(* IEC 61131-3 sources: plc-process-lib/tests/POUs/Suites/FB_ControlValve_Test, 43 files *)

(* ---- AutoSpNaNHoldsWithWarning.method.decl.st ---- *)
// Задание автоматики не число (NaN из Modbus/ПИД): выход удерживается, CV_WRN_SP_INVALID; конечное
// задание — снова к нему, предупреждение снято.
METHOD PRIVATE AutoSpNaNHoldsWithWarning
VAR
    fbTime   : FB_FakeTime;          // подменное время, старт 1 ч
    fbCv     : FB_ControlValve;      // клапан под тестом
    stCmd    : ST_ControlValveCmd;   // команды HMI
    stRetain : ST_DeviceRetain;      // режим Manual по умолчанию
    stCfg    : ST_ControlValveCfg;   // конфигурация (умолчания: 0…100 %, без рампы)
    uBits    : U_RealBits;           // NaN по битам
END_VAR

(* ---- AutoToManualBumpless.method.decl.st ---- *)
// Auto 70 %: задание Manual следит (70 %). Переход в Manual при задании автоматики 20 %: выход остаётся
// 70 %, xAutoActive = FALSE; задание оператора 60 % — рампа 5 %/с от 70 %: 65 % через 1 с.
METHOD PRIVATE AutoToManualBumpless
VAR
    fbTime   : FB_FakeTime;          // подменное время, старт 1 ч
    fbCv     : FB_ControlValve;      // клапан под тестом
    stCmd    : ST_ControlValveCmd;   // команды HMI
    stRetain : ST_DeviceRetain;      // режим Manual по умолчанию
    stCfg    : ST_ControlValveCfg;   // конфигурация (умолчания: 0…100 %, без рампы)
    iStep    : INT;                  // шаг цикла
END_VAR

(* ---- AutoToManualBumpless.method.impl.st ---- *)
coUnit.TEST('ControlValve_AutoToManual_Bumpless');

stRetain.eRemoteMode := E_DeviceMode.Auto;
fbCv.rPosSpAuto_pct := 70.0;
fbCv(itfTime := fbTime, stCmd := stCmd, stRetain := stRetain, stCfg := stCfg);
AssertEquals_REAL(Expected := 70.0, Actual := fbCv.rOut_pct, Delta := 0.0, Message := 'Auto 70 %');
AssertTrue(Condition := fbCv.xAutoActive, Message := 'xAutoActive');
AssertEquals_REAL(Expected := 70.0, Actual := stCmd.rPosSpMan_pct, Delta := 0.0,
                  Message := 'manual setpoint tracks in Auto');
stCfg.rRateUp_pctps := 5.0;
stCfg.rRateDown_pctps := 5.0;
stCmd.stCommon.xSetManual := TRUE;
fbCv.rPosSpAuto_pct := 20.0;
fbTime.Advance(tStep := T#100MS);
fbCv(itfTime := fbTime, stCmd := stCmd, stRetain := stRetain, stCfg := stCfg);
AssertTrue(Condition := fbCv.Mode = E_DeviceMode.Manual, Message := 'Manual');
AssertEquals_REAL(Expected := 70.0, Actual := fbCv.rOut_pct, Delta := 0.0, Message := 'no bump');
AssertFalse(Condition := fbCv.xAutoActive, Message := 'xAutoActive off in Manual');
stCmd.rPosSpMan_pct := 60.0;
FOR iStep := 1 TO 10 DO
    fbTime.Advance(tStep := T#100MS);
    fbCv(itfTime := fbTime, stCmd := stCmd, stRetain := stRetain, stCfg := stCfg);
END_FOR
// источник: tools/reference/valve_reference.py, сценарий cv_bumpless (70 -> 60, 5 %/s, 1.0 s)
AssertEquals_REAL(Expected := 65.0, Actual := fbCv.rOut_pct, Delta := 1.0E-4,
                  Message := 'ramp from 70 %: 65 % after 1 s');

coUnit.TEST_FINISHED();

(* ---- CfgChecksSetBits.method.decl.st ---- *)
// Каждая проверка CheckConfig даёт свой бит wCfgErr: пределы (min < 0, max > 100, min >= max), скорость
// (< 0, NaN), положение безопасности вне 0…100, рассогласование при подключённой ОС (допуск 0, tDev = 0;
// без ОС не проверяется), плотное закрытие (< 0, >= rOutMax), реакция на отказ вне перечисления,
// приоритет тревоги.
METHOD PRIVATE CfgChecksSetBits
VAR
    fbTime   : FB_FakeTime;          // подменное время, старт 1 ч
    fbCv     : FB_ControlValve;      // клапан под тестом
    stCmd    : ST_ControlValveCmd;   // команды HMI
    stRetain : ST_DeviceRetain;      // режим Manual по умолчанию
    stCfg    : ST_ControlValveCfg;   // конфигурация (умолчания: 0…100 %, без рампы)
    uBad     : U_TestValveEnum;      // значение вне перечисления
    uBits    : U_RealBits;           // NaN по битам
    stSlot   : ST_AlarmCfg;          // копия слота тревоги
END_VAR

(* ---- DefaultCfgPassesCheck.method.decl.st ---- *)
// Умолчания ST_ControlValveCfg проходят CheckConfig; тип ControlValve, слотов тревог 4, приоритеты по
// умолчанию (PositionerFault — Medium, InterlockAct — None); ток 4 мА при 0 %; Manual — xAutoActive нет.
METHOD PRIVATE DefaultCfgPassesCheck
VAR
    fbTime   : FB_FakeTime;          // подменное время, старт 1 ч
    fbCv     : FB_ControlValve;      // клапан под тестом
    stCmd    : ST_ControlValveCmd;   // команды HMI
    stRetain : ST_DeviceRetain;      // режим Manual по умолчанию
    stCfg    : ST_ControlValveCfg;   // конфигурация (умолчания: 0…100 %, без рампы)
    itfAlm   : I_Alarm;              // слот тревоги через интерфейс
END_VAR

(* ---- DeviationAsFaultGoesSafePosition.method.decl.st ---- *)
// Рассогласование — отказ (xDevIsFault), реакция SafePos (20 %), рампа 10 %/с, tDev = 5 с. Auto, выход
// 50 %, ОС 30 %: на 4 с отказа нет, на 5 с — CV_FLT_DEVIATION, Failure и сразу 20 % без рампы (бит
// SAFE_POS), xAutoActive = FALSE. Отказ фиксирован; Reset снимает, рампа к 50 % — от текущих 20 %.
METHOD PRIVATE DeviationAsFaultGoesSafePosition
VAR
    fbTime   : FB_FakeTime;          // подменное время, старт 1 ч
    fbCv     : FB_ControlValve;      // клапан под тестом
    stCmd    : ST_ControlValveCmd;   // команды HMI
    stRetain : ST_DeviceRetain;      // режим Manual по умолчанию
    stCfg    : ST_ControlValveCfg;   // конфигурация (умолчания: 0…100 %, без рампы)
    iStep    : INT;                  // шаг цикла
END_VAR

(* ---- DeviationAsFaultGoesSafePosition.method.impl.st ---- *)
coUnit.TEST('ControlValve_DeviationAsFault_GoesSafePosition');

stCfg.xFbUsed := TRUE;
stCfg.xDevIsFault := TRUE;
stCfg.eFaultAction := E_CvFaultAction.SafePos;
stCfg.rSafePos_pct := 20.0;
stCfg.tDev := T#5S;
stRetain.eRemoteMode := E_DeviceMode.Auto;
fbCv.rPosSpAuto_pct := 50.0;
fbCv.xPosFbValid := TRUE;
fbCv.rPosFb_pct := 50.0;
// Auto, 50 % (без рампы — сразу)
fbCv(itfTime := fbTime, stCmd := stCmd, stRetain := stRetain, stCfg := stCfg);
stCfg.rRateUp_pctps := 10.0;
stCfg.rRateDown_pctps := 10.0;
fbCv.rPosFb_pct := 30.0;
fbTime.Advance(tStep := T#1S);
// t1: клапан отстал
fbCv(itfTime := fbTime, stCmd := stCmd, stRetain := stRetain, stCfg := stCfg);
FOR iStep := 1 TO 4 DO                                                  // t1 + 4 с
    fbTime.Advance(tStep := T#1S);
    fbCv(itfTime := fbTime, stCmd := stCmd, stRetain := stRetain, stCfg := stCfg);
END_FOR
AssertEquals_WORD(Expected := 0, Actual := fbCv.stSts.stCommon.wFault, Message := 'no fault before tDev');
AssertEquals_REAL(Expected := 50.0, Actual := fbCv.rOut_pct, Delta := 0.0, Message := 'output 50 %');
fbTime.Advance(tStep := T#1S);
// t1 + 5 с
fbCv(itfTime := fbTime, stCmd := stCmd, stRetain := stRetain, stCfg := stCfg);
AssertEquals_WORD(Expected := GVL_Const.CV_FLT_DEVIATION, Actual := fbCv.stSts.stCommon.wFault,
                  Message := 'deviation fault');
AssertTrue(Condition := fbCv.Status = E_Ne107Status.Failure, Message := 'NE 107 Failure');
AssertEquals_REAL(Expected := 20.0, Actual := fbCv.rOut_pct, Delta := 0.0, Message := 'safe position at once, no ramp');
AssertEquals_WORD(Expected := GVL_Const.CV_STS_SAFE_POS,
                  Actual := fbCv.stSts.stCommon.wStatus AND GVL_Const.CV_STS_SAFE_POS, Message := 'SAFE_POS bit');
AssertFalse(Condition := fbCv.xAutoActive, Message := 'PID must track');
fbCv.rPosFb_pct := 20.0;
fbTime.Advance(tStep := T#1S);
fbCv(itfTime := fbTime, stCmd := stCmd, stRetain := stRetain, stCfg := stCfg);
AssertEquals_WORD(Expected := GVL_Const.CV_FLT_DEVIATION, Actual := fbCv.stSts.stCommon.wFault, Message := 'latched');
stCmd.stCommon.xReset := TRUE;
// без шага времени
fbCv(itfTime := fbTime, stCmd := stCmd, stRetain := stRetain, stCfg := stCfg);
AssertEquals_WORD(Expected := 0, Actual := fbCv.stSts.stCommon.wFault, Message := 'cleared by Reset');
AssertTrue(Condition := fbCv.stSts.stCommon.eCmdResult = E_CmdResult.Accepted, Message := 'Reset accepted');
AssertEquals_REAL(Expected := 20.0, Actual := fbCv.rOut_pct, Delta := 0.0,
                  Message := 'ramp starts from current output');
FOR iStep := 1 TO 10 DO
    fbTime.Advance(tStep := T#100MS);
    fbCv(itfTime := fbTime, stCmd := stCmd, stRetain := stRetain, stCfg := stCfg);
END_FOR
// источник: tools/reference/valve_reference.py, сценарий cv_return_ramp (20 -> 50, 10 %/s, 1.0 s)
AssertEquals_REAL(Expected := 30.0, Actual := fbCv.rOut_pct, Delta := 1.0E-4, Message := 'ramps back: 30 % after 1 s');
AssertTrue(Condition := fbCv.xAutoActive, Message := 'xAutoActive again');

coUnit.TEST_FINISHED();

(* ---- DeviationDuringRampIgnored.method.decl.st ---- *)
// Клапан не двигается (ОС 0 %), задание 0 -> 50 % с рампой 1 %/с (50 с): во время рампы рассогласование
// не контролируется. После конца рампы предупреждение — ровно через tDev = 10 с (на 9 с ещё нет).
METHOD PRIVATE DeviationDuringRampIgnored
VAR
    fbTime    : FB_FakeTime;          // подменное время, старт 1 ч
    fbCv      : FB_ControlValve;      // клапан под тестом
    stCmd     : ST_ControlValveCmd;   // команды HMI
    stRetain  : ST_DeviceRetain;      // режим Manual по умолчанию
    stCfg     : ST_ControlValveCfg;   // конфигурация (умолчания: 0…100 %, без рампы)
    iStep     : INT;                  // шаг цикла
    xEverWarn : BOOL;                 // предупреждение было во время рампы
END_VAR

(* ---- DeviationDuringRampIgnored.method.impl.st ---- *)
coUnit.TEST('ControlValve_DeviationDuringRamp_Ignored');

stCfg.xFbUsed := TRUE;
stCfg.tDev := T#10S;
stCfg.rRateUp_pctps := 1.0;
fbCv.xPosFbValid := TRUE;
fbCv.rPosFb_pct := 0.0;
// t0: задание 0
fbCv(itfTime := fbTime, stCmd := stCmd, stRetain := stRetain, stCfg := stCfg);
stCmd.rPosSpMan_pct := 50.0;
FOR iStep := 1 TO 50 DO                                                 // рампа 50 с
    fbTime.Advance(tStep := T#1S);
    fbCv(itfTime := fbTime, stCmd := stCmd, stRetain := stRetain, stCfg := stCfg);
    xEverWarn := xEverWarn OR (fbCv.stSts.stCommon.wWarning AND GVL_Const.CV_WRN_DEVIATION) <> 0;
END_FOR
AssertFalse(Condition := xEverWarn, Message := 'no deviation supervision while ramping');
AssertEquals_REAL(Expected := 50.0, Actual := fbCv.rOut_pct, Delta := 1.0E-4, Message := 'ramp finished at 50 %');
AssertEquals_WORD(Expected := 0, Actual := fbCv.stSts.stCommon.wStatus AND GVL_Const.CV_STS_RAMPING,
                  Message := 'RAMPING cleared');
FOR iStep := 1 TO 10 DO                                                 // 9 с после рампы
    fbTime.Advance(tStep := T#1S);
    fbCv(itfTime := fbTime, stCmd := stCmd, stRetain := stRetain, stCfg := stCfg);
END_FOR
AssertEquals_WORD(Expected := 0, Actual := fbCv.stSts.stCommon.wWarning AND GVL_Const.CV_WRN_DEVIATION,
                  Message := 'no warning before tDev after the ramp');
fbTime.Advance(tStep := T#1S);
fbCv(itfTime := fbTime, stCmd := stCmd, stRetain := stRetain, stCfg := stCfg);
AssertEquals_WORD(Expected := GVL_Const.CV_WRN_DEVIATION,
                  Actual := fbCv.stSts.stCommon.wWarning AND GVL_Const.CV_WRN_DEVIATION,
                  Message := 'deviation once the ramp ended and tDev passed');

coUnit.TEST_FINISHED();

(* ---- DeviationFaultResetStuckValveRetripsAfterTDev.method.decl.st ---- *)
// Рассогласование — отказ (xDevIsFault), реакция Hold, tDev = 5 с. Manual, задание 50 %, клапан
// заклинило на 30 %: на t0 + 5 с — CV_FLT_DEVIATION, выход удерживается (50 %), предупреждения
// рассогласования нет — это отказ. Reset при неснятой причине снимает отказ и начинает отсчёт tDev заново:
// на t1 + 4 с отказа нет, ровно на t1 + 5 с он возвращается.
METHOD PRIVATE DeviationFaultResetStuckValveRetripsAfterTDev
VAR
    fbTime   : FB_FakeTime;          // подменное время, старт 1 ч
    fbCv     : FB_ControlValve;      // клапан под тестом
    stCmd    : ST_ControlValveCmd;   // команды HMI
    stRetain : ST_DeviceRetain;      // режим Manual по умолчанию
    stCfg    : ST_ControlValveCfg;   // конфигурация (умолчания: 0…100 %, без рампы, Hold)
    iStep    : INT;                  // шаг цикла
END_VAR

(* ---- DeviationFaultResetStuckValveRetripsAfterTDev.method.impl.st ---- *)
coUnit.TEST('ControlValve_DeviationFaultReset_StuckValveRetripsAfterTDev');

stCfg.xFbUsed := TRUE;
stCfg.xDevIsFault := TRUE;
stCfg.tDev := T#5S;
stCmd.rPosSpMan_pct := 50.0;
fbCv.xPosFbValid := TRUE;
fbCv.rPosFb_pct := 30.0;
// выход 50 %, клапан стоит на 30 %
fbCv(itfTime := fbTime, stCmd := stCmd, stRetain := stRetain, stCfg := stCfg);
// t0: первый вызов, в котором оценивается рассогласование (выход уже подан)
fbCv(itfTime := fbTime, stCmd := stCmd, stRetain := stRetain, stCfg := stCfg);
FOR iStep := 1 TO 5 DO                                                  // t0 + 5 с
    fbTime.Advance(tStep := T#1S);
    fbCv(itfTime := fbTime, stCmd := stCmd, stRetain := stRetain, stCfg := stCfg);
END_FOR
AssertEquals_WORD(Expected := GVL_Const.CV_FLT_DEVIATION, Actual := fbCv.stSts.stCommon.wFault,
                  Message := 'deviation fault');
AssertEquals_WORD(Expected := 0, Actual := fbCv.stSts.stCommon.wWarning AND GVL_Const.CV_WRN_DEVIATION,
                  Message := 'fault, not warning');
AssertEquals_REAL(Expected := 50.0, Actual := fbCv.rOut_pct, Delta := 0.0, Message := 'Hold keeps the output');
stCmd.stCommon.xReset := TRUE;
// t1: Reset, клапан всё так же на 30 %
fbCv(itfTime := fbTime, stCmd := stCmd, stRetain := stRetain, stCfg := stCfg);
AssertEquals_WORD(Expected := 0, Actual := fbCv.stSts.stCommon.wFault, Message := 'cleared by Reset');
FOR iStep := 1 TO 4 DO                                                  // t1 + 4 с
    fbTime.Advance(tStep := T#1S);
    fbCv(itfTime := fbTime, stCmd := stCmd, stRetain := stRetain, stCfg := stCfg);
END_FOR
AssertEquals_WORD(Expected := 0, Actual := fbCv.stSts.stCommon.wFault, Message := 'tDev restarted by Reset');
fbTime.Advance(tStep := T#1S);
// t1 + 5 с
fbCv(itfTime := fbTime, stCmd := stCmd, stRetain := stRetain, stCfg := stCfg);
AssertEquals_WORD(Expected := GVL_Const.CV_FLT_DEVIATION, Actual := fbCv.stSts.stCommon.wFault,
                  Message := 'stuck valve trips again after tDev');

coUnit.TEST_FINISHED();

(* ---- DeviationWarningAfterDelay.method.decl.st ---- *)
// ОС подключена, допуск 5 %, tDev = 30 с. Выход 50 %, ОС 40 %: до 29 с предупреждения нет, ровно на 30 с —
// CV_WRN_DEVIATION, NE 107 OutOfSpecification, тревога слота Deviation; отказа нет, выход не меняется,
// rDeviation_pct = 10 %. ОС 48 % — предупреждение снято, бит AT_SETPOINT.
METHOD PRIVATE DeviationWarningAfterDelay
VAR
    fbTime   : FB_FakeTime;          // подменное время, старт 1 ч
    fbCv     : FB_ControlValve;      // клапан под тестом
    stCmd    : ST_ControlValveCmd;   // команды HMI
    stRetain : ST_DeviceRetain;      // режим Manual по умолчанию
    stCfg    : ST_ControlValveCfg;   // конфигурация (умолчания: 0…100 %, без рампы)
    iStep    : INT;                  // шаг цикла
    itfAlm   : I_Alarm;              // слот тревоги через интерфейс
END_VAR

(* ---- DeviationWarningAfterDelay.method.impl.st ---- *)
coUnit.TEST('ControlValve_Deviation_WarningAfterDelay');

stCfg.xFbUsed := TRUE;
stCmd.rPosSpMan_pct := 50.0;
fbCv.xPosFbValid := TRUE;
fbCv.rPosFb_pct := 50.0;
// на задании
fbCv(itfTime := fbTime, stCmd := stCmd, stRetain := stRetain, stCfg := stCfg);
AssertEquals_WORD(Expected := GVL_Const.CV_STS_AT_SETPOINT,
                  Actual := fbCv.stSts.stCommon.wStatus AND GVL_Const.CV_STS_AT_SETPOINT, Message := 'AT_SETPOINT');
fbCv.rPosFb_pct := 40.0;
fbTime.Advance(tStep := T#1S);
// t1: рассогласование 10 %
fbCv(itfTime := fbTime, stCmd := stCmd, stRetain := stRetain, stCfg := stCfg);
FOR iStep := 1 TO 29 DO                                                 // t1 + 29 с
    fbTime.Advance(tStep := T#1S);
    fbCv(itfTime := fbTime, stCmd := stCmd, stRetain := stRetain, stCfg := stCfg);
END_FOR
AssertEquals_WORD(Expected := 0, Actual := fbCv.stSts.stCommon.wWarning AND GVL_Const.CV_WRN_DEVIATION,
                  Message := 'no warning before tDev');
fbTime.Advance(tStep := T#1S);
// t1 + 30 с
fbCv(itfTime := fbTime, stCmd := stCmd, stRetain := stRetain, stCfg := stCfg);
AssertEquals_WORD(Expected := GVL_Const.CV_WRN_DEVIATION,
                  Actual := fbCv.stSts.stCommon.wWarning AND GVL_Const.CV_WRN_DEVIATION,
Message := 'deviation warning');
AssertTrue(Condition := fbCv.Status = E_Ne107Status.OutOfSpecification, Message := 'NE 107 OutOfSpecification');
AssertEquals_WORD(Expected := 0, Actual := fbCv.stSts.stCommon.wFault, Message := 'warning, not fault');
AssertEquals_REAL(Expected := 50.0, Actual := fbCv.rOut_pct, Delta := 0.0, Message := 'control continues');
AssertEquals_REAL(Expected := 10.0, Actual := fbCv.stSts.rDeviation_pct, Delta := 1.0E-5, Message := 'deviation 10 %');
AssertEquals_WORD(Expected := 0, Actual := fbCv.stSts.stCommon.wStatus AND GVL_Const.CV_STS_AT_SETPOINT,
                  Message := 'not at setpoint');
itfAlm := fbCv.GetAlarm(uiIndex := E_CvAlarm.Deviation);
AssertTrue(Condition := itfAlm.Active, Message := 'Deviation alarm active');
fbCv.rPosFb_pct := 48.0;
fbTime.Advance(tStep := T#1S);
fbCv(itfTime := fbTime, stCmd := stCmd, stRetain := stRetain, stCfg := stCfg);
AssertEquals_WORD(Expected := 0, Actual := fbCv.stSts.stCommon.wWarning AND GVL_Const.CV_WRN_DEVIATION,
                  Message := 'warning clears within tolerance');
AssertEquals_WORD(Expected := GVL_Const.CV_STS_AT_SETPOINT,
                  Actual := fbCv.stSts.stCommon.wStatus AND GVL_Const.CV_STS_AT_SETPOINT,
Message := 'AT_SETPOINT again');
AssertTrue(Condition := fbCv.Status = E_Ne107Status.Good, Message := 'NE 107 Good');

coUnit.TEST_FINISHED();

(* ---- FbInvalidMaintenanceRequiredKeepsControl.method.decl.st ---- *)
// ОС подключена, но недостоверна: CV_WRN_FB_INVALID, NE 107 MaintenanceRequired, тревога FbFailure;
// клапан управляется (30 % -> 60 %), xAutoActive и Available; рассогласование без ОС не контролируется
// дольше tDev. NaN при признаке «достоверна» — тоже отказ ОС.
METHOD PRIVATE FbInvalidMaintenanceRequiredKeepsControl
VAR
    fbTime   : FB_FakeTime;          // подменное время, старт 1 ч
    fbCv     : FB_ControlValve;      // клапан под тестом
    stCmd    : ST_ControlValveCmd;   // команды HMI
    stRetain : ST_DeviceRetain;      // режим Manual по умолчанию
    stCfg    : ST_ControlValveCfg;   // конфигурация (умолчания: 0…100 %, без рампы)
    iStep    : INT;                  // шаг цикла
    itfAlm   : I_Alarm;              // слот тревоги через интерфейс
    uBits    : U_RealBits;           // NaN по битам
END_VAR

(* ---- FbInvalidMaintenanceRequiredKeepsControl.method.impl.st ---- *)
coUnit.TEST('ControlValve_FbInvalid_MaintenanceRequiredKeepsControl');

stCfg.xFbUsed := TRUE;
stCfg.tDev := T#5S;
stRetain.eRemoteMode := E_DeviceMode.Auto;
fbCv.rPosSpAuto_pct := 30.0;
fbCv.xPosFbValid := FALSE;
fbCv(itfTime := fbTime, stCmd := stCmd, stRetain := stRetain, stCfg := stCfg);
AssertEquals_WORD(Expected := GVL_Const.CV_WRN_FB_INVALID, Actual := fbCv.stSts.stCommon.wWarning,
                  Message := 'FB_INVALID');
AssertTrue(Condition := fbCv.Status = E_Ne107Status.MaintenanceRequired, Message := 'NE 107 MaintenanceRequired');
AssertEquals_REAL(Expected := 30.0, Actual := fbCv.rOut_pct, Delta := 0.0, Message := 'control continues');
AssertTrue(Condition := fbCv.xAutoActive, Message := 'xAutoActive');
AssertTrue(Condition := fbCv.Available, Message := 'available');
itfAlm := fbCv.GetAlarm(uiIndex := E_CvAlarm.FbFailure);
AssertTrue(Condition := itfAlm.Active, Message := 'FbFailure alarm');
FOR iStep := 1 TO 10 DO                                                 // дольше tDev
    fbTime.Advance(tStep := T#1S);
    fbCv(itfTime := fbTime, stCmd := stCmd, stRetain := stRetain, stCfg := stCfg);
END_FOR
AssertEquals_WORD(Expected := 0, Actual := fbCv.stSts.stCommon.wWarning AND GVL_Const.CV_WRN_DEVIATION,
                  Message := 'no deviation supervision without feedback');
AssertEquals_WORD(Expected := 0, Actual := fbCv.stSts.stCommon.wFault, Message := 'no fault');
fbCv.rPosSpAuto_pct := 60.0;
fbTime.Advance(tStep := T#100MS);
fbCv(itfTime := fbTime, stCmd := stCmd, stRetain := stRetain, stCfg := stCfg);
AssertEquals_REAL(Expected := 60.0, Actual := fbCv.rOut_pct, Delta := 0.0, Message := 'follows new setpoint');
uBits.dwValue := 16#7FC00000;
fbCv.rPosFb_pct := uBits.rValue;
fbCv.xPosFbValid := TRUE;
fbTime.Advance(tStep := T#100MS);
fbCv(itfTime := fbTime, stCmd := stCmd, stRetain := stRetain, stCfg := stCfg);
AssertEquals_WORD(Expected := GVL_Const.CV_WRN_FB_INVALID,
                  Actual := fbCv.stSts.stCommon.wWarning AND GVL_Const.CV_WRN_FB_INVALID,
                  Message := 'NaN feedback invalid');
// AssertEquals_REAL пропускает NaN (ABS(NaN) > Delta = FALSE): конечность проверяется отдельно
AssertTrue(Condition := F_IsFinite(rIn := fbCv.rOut_pct) AND F_IsFinite(rIn := fbCv.rOut_mA),
           Message := 'output finite with NaN feedback');
AssertTrue(Condition := F_IsFinite(rIn := fbCv.stSts.rDeviation_pct), Message := 'deviation finite');
AssertEquals_REAL(Expected := 0.0, Actual := fbCv.stSts.rDeviation_pct, Delta := 0.0,
                  Message := 'no deviation without valid feedback (CV-8)');
AssertEquals_REAL(Expected := 60.0, Actual := fbCv.rOut_pct, Delta := 0.0, Message := 'control continues');

coUnit.TEST_FINISHED();

(* ---- FbNaNEventAndStsFinite.method.decl.st ---- *)
// ОС положения NaN при xPosFbValid = TRUE (мусор Modbus): тревога FbFailure; значение её события и stSts.rPosFb_pct
// конечны — 0.0 (R6: журнал и карта регистров NaN не получают), рассогласование 0, выход удерживается.
METHOD PRIVATE FbNaNEventAndStsFinite
VAR
    fbTime   : FB_FakeTime;          // подменное время, старт 1 ч
    fbCv     : FB_ControlValve;      // клапан под тестом
    stCmd    : ST_ControlValveCmd;   // команды HMI
    stRetain : ST_DeviceRetain;      // режим Manual по умолчанию
    stCfg    : ST_ControlValveCfg;   // конфигурация (умолчания: 0…100 %, без рампы)

    fbSink   : FB_TestSink;          // приёмник событий
    stEv     : ST_AlarmEvent;        // последнее событие
    uBits    : U_RealBits;           // NaN по битам
END_VAR

(* ---- InterlockFirstOutKeptUntilResetOrOos.method.decl.st ---- *)
// Первопричина держится (CV-9): блокировка бит 2, затем добавился бит 0 (16#0005) — uiFirstOut = 2 не меняется.
// Reset снимает её; пока слово блокировок не 0, новой первопричины нет. Слово вернулось в 0, затем бит 1 —
// первопричина 1; вход в OutOfService её снимает.
METHOD PRIVATE InterlockFirstOutKeptUntilResetOrOos
VAR
    fbTime   : FB_FakeTime;          // подменное время, старт 1 ч
    fbCv     : FB_ControlValve;      // клапан под тестом
    stCmd    : ST_ControlValveCmd;   // команды HMI
    stRetain : ST_DeviceRetain;      // режим Manual по умолчанию
    stCfg    : ST_ControlValveCfg;   // конфигурация (умолчания: 0…100 %, без рампы)
END_VAR

(* ---- InterlockInManualStaysAtSafePosition.method.decl.st ---- *)
// Manual, задание оператора 70 %. Блокировка: выход сразу в положение безопасности 15 %, задание
// Manual следит за ним (оператор не управляет выходом). Блокировка снята: Manual остаётся в 15 % —
// клапан сам к прежнему заданию оператора не уходит (CV-6, как у FB_Valve и двигателя).
METHOD PRIVATE InterlockInManualStaysAtSafePosition
VAR
    fbTime   : FB_FakeTime;          // подменное время, старт 1 ч
    fbCv     : FB_ControlValve;      // клапан под тестом
    stCmd    : ST_ControlValveCmd;   // команды HMI
    stRetain : ST_DeviceRetain;      // режим Manual по умолчанию
    stCfg    : ST_ControlValveCfg;   // конфигурация (умолчания: 0…100 %, без рампы)
END_VAR

(* ---- InterlockSafePosBypassesRamp.method.decl.st ---- *)
// Блокировка (бит 2) при рампе 1 %/с: выход 60 % -> 10 % в том же вызове, мимо рампы и ниже rOutMin
// (20 %); биты SAFE_POS и INTERLOCKED, wInterlock, первопричина 2; xAutoActive = FALSE; задание Manual
// следит за принудительным выходом. После снятия — рампа от 10 %: 11 % через 1 с.
METHOD PRIVATE InterlockSafePosBypassesRamp
VAR
    fbTime   : FB_FakeTime;          // подменное время, старт 1 ч
    fbCv     : FB_ControlValve;      // клапан под тестом
    stCmd    : ST_ControlValveCmd;   // команды HMI
    stRetain : ST_DeviceRetain;      // режим Manual по умолчанию
    stCfg    : ST_ControlValveCfg;   // конфигурация (умолчания: 0…100 %, без рампы)
END_VAR

(* ---- InvalidCfgAtRuntimeKeepsLastValid.method.decl.st ---- *)
// Cfg испорчена в работе (скорость < 0): бит CV_CFG_RATE и CheckFunction, рампа продолжается по
// последней корректной Cfg (10 %/с): 10 % через 1 с.
METHOD PRIVATE InvalidCfgAtRuntimeKeepsLastValid
VAR
    fbTime   : FB_FakeTime;          // подменное время, старт 1 ч
    fbCv     : FB_ControlValve;      // клапан под тестом
    stCmd    : ST_ControlValveCmd;   // команды HMI
    stRetain : ST_DeviceRetain;      // режим Manual по умолчанию
    stCfg    : ST_ControlValveCfg;   // конфигурация (умолчания: 0…100 %, без рампы)
    iStep    : INT;                  // шаг цикла
END_VAR

(* ---- InvalidCfgAtRuntimeKeepsLastValid.method.impl.st ---- *)
coUnit.TEST('ControlValve_InvalidCfgAtRuntime_KeepsLastValid');

stCfg.rRateUp_pctps := 10.0;
fbCv(itfTime := fbTime, stCmd := stCmd, stRetain := stRetain, stCfg := stCfg);
stCmd.rPosSpMan_pct := 50.0;
stCfg.rRateUp_pctps := -1.0;
FOR iStep := 1 TO 10 DO
    fbTime.Advance(tStep := T#100MS);
    fbCv(itfTime := fbTime, stCmd := stCmd, stRetain := stRetain, stCfg := stCfg);
END_FOR
AssertEquals_WORD(Expected := GVL_Const.CV_CFG_RATE, Actual := fbCv.stSts.stCommon.wCfgErr, Message := 'CV_CFG_RATE');
AssertTrue(Condition := fbCv.Status = E_Ne107Status.CheckFunction, Message := 'NE 107 CheckFunction');
// источник: tools/reference/valve_reference.py, сценарий cv_manual_ramp (up 1.0 s)
AssertEquals_REAL(Expected := 10.0, Actual := fbCv.rOut_pct, Delta := 1.0E-4, Message := 'ramp with last valid rate');

coUnit.TEST_FINISHED();

(* ---- InvalidCfgStartupSafePosition.method.decl.st ---- *)
// Корректной Cfg ещё не было (rOutMin >= rOutMax): CV_CFG_LIMITS, CheckFunction; выход — положение
// безопасности из поданной Cfg (30 %, 8,8 мА) и в Auto, xAutoActive = FALSE, задание Manual следит.
// Положение безопасности NaN — 0 % (4 мА), 150 % — ограничено 100 %.
METHOD PRIVATE InvalidCfgStartupSafePosition
VAR
    fbTime      : FB_FakeTime;          // подменное время
    fbCv        : FB_ControlValve;      // клапан с неверными пределами
    fbCvBad     : FB_ControlValve;      // клапан с неверным положением безопасности
    stCmd       : ST_ControlValveCmd;   // команды
    stCmdBad    : ST_ControlValveCmd;   // команды второго клапана
    stRetain    : ST_DeviceRetain;      // режим
    stRetainBad : ST_DeviceRetain;      // режим второго клапана
    stCfg       : ST_ControlValveCfg;   // rOutMin >= rOutMax
    stCfgBad    : ST_ControlValveCfg;   // rSafePos_pct вне 0…100
    uBits       : U_RealBits;           // NaN по битам
    iStep       : INT;                  // шаг цикла
END_VAR

(* ---- InvalidCfgStartupSafePosition.method.impl.st ---- *)
coUnit.TEST('ControlValve_InvalidCfg_StartupSafePosition');

stCfg.rOutMin_pct := 50.0;
stCfg.rOutMax_pct := 40.0;
stCfg.rSafePos_pct := 30.0;
stRetain.eRemoteMode := E_DeviceMode.Auto;
fbCv.rPosSpAuto_pct := 70.0;
fbCv(itfTime := fbTime, stCmd := stCmd, stRetain := stRetain, stCfg := stCfg);
AssertEquals_WORD(Expected := GVL_Const.CV_CFG_LIMITS, Actual := fbCv.stSts.stCommon.wCfgErr,
                  Message := 'CV_CFG_LIMITS');
AssertTrue(Condition := fbCv.Status = E_Ne107Status.CheckFunction, Message := 'NE 107 CheckFunction');
AssertEquals_REAL(Expected := 30.0, Actual := fbCv.rOut_pct, Delta := 0.0, Message := 'safe position from cfg');
// источник: tools/reference/valve_reference.py, сценарий cv_ma (30 %)
AssertEquals_REAL(Expected := 8.8, Actual := fbCv.rOut_mA, Delta := 1.0E-5, Message := '30 % = 8.8 mA');
AssertEquals_WORD(Expected := GVL_Const.CV_STS_SAFE_POS,
                  Actual := fbCv.stSts.stCommon.wStatus AND GVL_Const.CV_STS_SAFE_POS, Message := 'SAFE_POS');
AssertFalse(Condition := fbCv.xAutoActive, Message := 'no xAutoActive without valid cfg');
AssertFalse(Condition := fbCv.Available, Message := 'not available');
AssertEquals_REAL(Expected := 30.0, Actual := stCmd.rPosSpMan_pct, Delta := 0.0, Message := 'manual setpoint tracks');
FOR iStep := 1 TO 10 DO
    fbTime.Advance(tStep := T#100MS);
    fbCv(itfTime := fbTime, stCmd := stCmd, stRetain := stRetain, stCfg := stCfg);
END_FOR
AssertEquals_REAL(Expected := 30.0, Actual := fbCv.rOut_pct, Delta := 0.0, Message := 'stays at safe position');
uBits.dwValue := 16#7FC00000;
stCfgBad.rSafePos_pct := uBits.rValue;
fbCvBad(itfTime := fbTime, stCmd := stCmdBad, stRetain := stRetainBad, stCfg := stCfgBad);
AssertEquals_WORD(Expected := GVL_Const.CV_CFG_SAFE_POS, Actual := fbCvBad.stSts.stCommon.wCfgErr,
                  Message := 'CV_CFG_SAFE_POS');
// AssertEquals_REAL пропускает NaN (ABS(NaN) > Delta = FALSE): конечность проверяется отдельно
AssertTrue(Condition := F_IsFinite(rIn := fbCvBad.rOut_pct) AND F_IsFinite(rIn := fbCvBad.rOut_mA),
           Message := 'NaN safe position: output finite');
AssertTrue(Condition := F_IsFinite(rIn := stCmdBad.rPosSpMan_pct), Message := 'manual setpoint tracking finite');
AssertEquals_REAL(Expected := 0.0, Actual := fbCvBad.rOut_pct, Delta := 0.0, Message := 'NaN safe position: 0 %');
AssertEquals_REAL(Expected := 4.0, Actual := fbCvBad.rOut_mA, Delta := 1.0E-5, Message := '4 mA');
stCfgBad.rSafePos_pct := 150.0;
fbTime.Advance(tStep := T#100MS);
fbCvBad(itfTime := fbTime, stCmd := stCmdBad, stRetain := stRetainBad, stCfg := stCfgBad);
AssertEquals_REAL(Expected := 100.0, Actual := fbCvBad.rOut_pct, Delta := 0.0, Message := 'limited to 100 %');

coUnit.TEST_FINISHED();

(* ---- Invert20mAAtZero.method.decl.st ---- *)
// Инверсия выхода: 0 % — 20 мА, 25 % — 16 мА, 100 % — 4 мА; без инверсии 25 % — 8 мА. Ток — и в выходе,
// и в Sts.
METHOD PRIVATE Invert20mAAtZero
VAR
    fbTime   : FB_FakeTime;          // подменное время, старт 1 ч
    fbCv     : FB_ControlValve;      // клапан под тестом
    stCmd    : ST_ControlValveCmd;   // команды HMI
    stRetain : ST_DeviceRetain;      // режим Manual по умолчанию
    stCfg    : ST_ControlValveCfg;   // конфигурация (умолчания: 0…100 %, без рампы)
END_VAR

(* ---- LocalFeedbackOutOfRangeOutputClamped.method.decl.st ---- *)
// Local: выход следует ОС, но только в пределах хода 0…100 %. Датчик положения на закрытом клапане
// показывает чуть ниже нуля (-1,5 %, сигнал ещё достоверен): выход 0 % и 4,0 мА, а не 3,76 мА — ток ниже
// 4 мА позиционер с питанием от токовой петли может не держать (минимальный ток — по паспорту
// позиционера). ОС 102,5 % — выход 100 % и 20,0 мА, а не 20,4 мА. С инверсией: 100 % — 4,0 мА, -1,5 % —
// 20,0 мА. Возврат в Manual — без рывка от ограниченного выхода.
METHOD PRIVATE LocalFeedbackOutOfRangeOutputClamped
VAR
    fbTime   : FB_FakeTime;          // подменное время, старт 1 ч
    fbCv     : FB_ControlValve;      // клапан под тестом
    stCmd    : ST_ControlValveCmd;   // команды HMI
    stRetain : ST_DeviceRetain;      // режим Manual по умолчанию
    stCfg    : ST_ControlValveCfg;   // конфигурация (умолчания: 0…100 %, без рампы)
END_VAR

(* ---- LocalTracksFeedback.method.decl.st ---- *)
// Local (позиционер на месте): выход сразу следует ОС 37 % без рампы, задание Manual тоже; ОС
// недостоверна — удержание и CV_WRN_FB_INVALID; ОС 42 % — 42 %. Возврат в Manual — без рывка.
METHOD PRIVATE LocalTracksFeedback
VAR
    fbTime   : FB_FakeTime;          // подменное время, старт 1 ч
    fbCv     : FB_ControlValve;      // клапан под тестом
    stCmd    : ST_ControlValveCmd;   // команды HMI
    stRetain : ST_DeviceRetain;      // режим Manual по умолчанию
    stCfg    : ST_ControlValveCfg;   // конфигурация (умолчания: 0…100 %, без рампы)
END_VAR

(* ---- ManualSetpointRateLimited.method.decl.st ---- *)
// Manual, рост 10 %/с, спад 20 %/с, шаг 0,1 с. Задание 0 -> 50 %: 10 % через 1 с, 49 % на 4,9 с, 50 % на
// 5,0 с (бит RAMPING снят); задание 50 -> 10 %: 30 % через 1 с, 10 % через 2 с. Задание оператора в
// Manual ФБ не переписывает.
METHOD PRIVATE ManualSetpointRateLimited
VAR
    fbTime   : FB_FakeTime;          // подменное время, старт 1 ч
    fbCv     : FB_ControlValve;      // клапан под тестом
    stCmd    : ST_ControlValveCmd;   // команды HMI
    stRetain : ST_DeviceRetain;      // режим Manual по умолчанию
    stCfg    : ST_ControlValveCfg;   // конфигурация (умолчания: 0…100 %, без рампы)
    iStep    : INT;                  // шаг цикла
END_VAR

(* ---- ManualSetpointRateLimited.method.impl.st ---- *)
coUnit.TEST('ControlValve_ManualSetpoint_RateLimited');

stCfg.rRateUp_pctps := 10.0;
stCfg.rRateDown_pctps := 20.0;
// t0: задание 0
fbCv(itfTime := fbTime, stCmd := stCmd, stRetain := stRetain, stCfg := stCfg);
stCmd.rPosSpMan_pct := 50.0;
FOR iStep := 1 TO 10 DO                                                 // t0 + 1,0 с
    fbTime.Advance(tStep := T#100MS);
    fbCv(itfTime := fbTime, stCmd := stCmd, stRetain := stRetain, stCfg := stCfg);
END_FOR
// источник: tools/reference/valve_reference.py, сценарий cv_manual_ramp (up 1.0 s)
AssertEquals_REAL(Expected := 10.0, Actual := fbCv.rOut_pct, Delta := 1.0E-4, Message := '10 % after 1 s');
AssertEquals_REAL(Expected := 50.0, Actual := fbCv.stSts.rPosSp_pct, Delta := 0.0, Message := 'setpoint before ramp');
AssertEquals_WORD(Expected := GVL_Const.CV_STS_RAMPING,
                  Actual := fbCv.stSts.stCommon.wStatus AND GVL_Const.CV_STS_RAMPING, Message := 'RAMPING bit');
AssertEquals_REAL(Expected := 50.0, Actual := stCmd.rPosSpMan_pct, Delta := 0.0,
                  Message := 'operator setpoint kept in Manual');
FOR iStep := 11 TO 49 DO                                                // t0 + 4,9 с
    fbTime.Advance(tStep := T#100MS);
    fbCv(itfTime := fbTime, stCmd := stCmd, stRetain := stRetain, stCfg := stCfg);
END_FOR
// источник: tools/reference/valve_reference.py, сценарий cv_manual_ramp (up 4.9 s)
AssertEquals_REAL(Expected := 49.0, Actual := fbCv.rOut_pct, Delta := 1.0E-4, Message := '49 % at 4.9 s');
fbTime.Advance(tStep := T#100MS);
// t0 + 5,0 с
fbCv(itfTime := fbTime, stCmd := stCmd, stRetain := stRetain, stCfg := stCfg);
// источник: tools/reference/valve_reference.py, сценарий cv_manual_ramp (up 5.0 s)
AssertEquals_REAL(Expected := 50.0, Actual := fbCv.rOut_pct, Delta := 1.0E-4, Message := '50 % at 5.0 s');
AssertEquals_WORD(Expected := 0, Actual := fbCv.stSts.stCommon.wStatus AND GVL_Const.CV_STS_RAMPING,
                  Message := 'ramp finished');
stCmd.rPosSpMan_pct := 10.0;
FOR iStep := 1 TO 10 DO
    fbTime.Advance(tStep := T#100MS);
    fbCv(itfTime := fbTime, stCmd := stCmd, stRetain := stRetain, stCfg := stCfg);
END_FOR
// источник: tools/reference/valve_reference.py, сценарий cv_manual_ramp (down 1.0 s)
AssertEquals_REAL(Expected := 30.0, Actual := fbCv.rOut_pct, Delta := 1.0E-4, Message := 'down 20 %/s: 30 % after 1 s');
FOR iStep := 11 TO 20 DO
    fbTime.Advance(tStep := T#100MS);
    fbCv(itfTime := fbTime, stCmd := stCmd, stRetain := stRetain, stCfg := stCfg);
END_FOR
// источник: tools/reference/valve_reference.py, сценарий cv_manual_ramp (down 2.0 s, mA at 10 %)
AssertEquals_REAL(Expected := 10.0, Actual := fbCv.rOut_pct, Delta := 1.0E-4, Message := '10 % after 2 s');
AssertEquals_REAL(Expected := 5.6, Actual := fbCv.rOut_mA, Delta := 1.0E-4, Message := '10 % = 5.6 mA');

coUnit.TEST_FINISHED();

(* ---- OosEntryClearsLatchedDeviation.method.decl.st ---- *)
// Зафиксированный отказ рассогласования снимается входом в OutOfService; после выхода в Manual отказа
// нет.
METHOD PRIVATE OosEntryClearsLatchedDeviation
VAR
    fbTime   : FB_FakeTime;          // подменное время, старт 1 ч
    fbCv     : FB_ControlValve;      // клапан под тестом
    stCmd    : ST_ControlValveCmd;   // команды HMI
    stRetain : ST_DeviceRetain;      // режим Manual по умолчанию
    stCfg    : ST_ControlValveCfg;   // конфигурация (умолчания: 0…100 %, без рампы)
    iStep    : INT;                  // шаг цикла
END_VAR

(* ---- OosEntryClearsLatchedDeviation.method.impl.st ---- *)
coUnit.TEST('ControlValve_OosEntry_ClearsLatchedDeviation');

stCfg.xFbUsed := TRUE;
stCfg.xDevIsFault := TRUE;
stCfg.tDev := T#2S;
stCmd.rPosSpMan_pct := 50.0;
fbCv.xPosFbValid := TRUE;
fbCv.rPosFb_pct := 10.0;
fbCv(itfTime := fbTime, stCmd := stCmd, stRetain := stRetain, stCfg := stCfg);
FOR iStep := 1 TO 3 DO
    fbTime.Advance(tStep := T#1S);
    fbCv(itfTime := fbTime, stCmd := stCmd, stRetain := stRetain, stCfg := stCfg);
END_FOR
AssertEquals_WORD(Expected := GVL_Const.CV_FLT_DEVIATION, Actual := fbCv.stSts.stCommon.wFault, Message := 'latched');
stCmd.stCommon.xSetOos := TRUE;
fbTime.Advance(tStep := T#100MS);
fbCv(itfTime := fbTime, stCmd := stCmd, stRetain := stRetain, stCfg := stCfg);
AssertTrue(Condition := fbCv.Mode = E_DeviceMode.OutOfService, Message := 'OutOfService');
AssertEquals_WORD(Expected := 0, Actual := fbCv.stSts.stCommon.wFault, Message := 'OOS entry clears the latch');
stCmd.stCommon.xSetManual := TRUE;
fbCv.rPosFb_pct := 50.0;
fbTime.Advance(tStep := T#100MS);
fbCv(itfTime := fbTime, stCmd := stCmd, stRetain := stRetain, stCfg := stCfg);
AssertTrue(Condition := fbCv.Mode = E_DeviceMode.Manual, Message := 'Manual');
AssertEquals_WORD(Expected := 0, Actual := fbCv.stSts.stCommon.wFault, Message := 'no fault after OOS');

coUnit.TEST_FINISHED();

(* ---- OutOfServiceHoldsOutput.method.decl.st ---- *)
// OutOfService: выход удерживается (40 %), задание, блокировка и отказ позиционера не действуют, задание
// Manual следит за удерживаемым выходом, NE 107 CheckFunction.
METHOD PRIVATE OutOfServiceHoldsOutput
VAR
    fbTime   : FB_FakeTime;          // подменное время, старт 1 ч
    fbCv     : FB_ControlValve;      // клапан под тестом
    stCmd    : ST_ControlValveCmd;   // команды HMI
    stRetain : ST_DeviceRetain;      // режим Manual по умолчанию
    stCfg    : ST_ControlValveCfg;   // конфигурация (умолчания: 0…100 %, без рампы)
END_VAR

(* ---- OutputLimitsClamp.method.decl.st ---- *)
// Пределы 10…90 %: задание Manual 95 % — выход 90 % (бит LIMITED_MAX), 5 % — 10 % (LIMITED_MIN); в Auto
// 120 % — 90 %, 55 % — без ограничения. rPosSp_pct — задание после пределов.
METHOD PRIVATE OutputLimitsClamp
VAR
    fbTime   : FB_FakeTime;          // подменное время, старт 1 ч
    fbCv     : FB_ControlValve;      // клапан под тестом
    stCmd    : ST_ControlValveCmd;   // команды HMI
    stRetain : ST_DeviceRetain;      // режим Manual по умолчанию
    stCfg    : ST_ControlValveCfg;   // конфигурация (умолчания: 0…100 %, без рампы)
    wLimBits : WORD;                 // биты LIMITED_MIN и LIMITED_MAX
END_VAR

(* ---- PositionerFaultHoldAction.method.decl.st ---- *)
// Отказ позиционера с реакцией Hold (по умолчанию): выход удерживается (40 %) при смене задания, бита
// SAFE_POS нет; отказ ушёл — выход к заданию 70 %.
METHOD PRIVATE PositionerFaultHoldAction
VAR
    fbTime   : FB_FakeTime;          // подменное время, старт 1 ч
    fbCv     : FB_ControlValve;      // клапан под тестом
    stCmd    : ST_ControlValveCmd;   // команды HMI
    stRetain : ST_DeviceRetain;      // режим Manual по умолчанию
    stCfg    : ST_ControlValveCfg;   // конфигурация (умолчания: 0…100 %, без рампы)
END_VAR

(* ---- PositionerFaultSafePosAction.method.decl.st ---- *)
// Отказ позиционера, реакция SafePos (100 %, «открыть при отказе»), рампа 2 %/с: выход 40 % -> 100 % в
// том же вызове, CV_FLT_POSITIONER, Failure, SAFE_POS. Отказ не фиксируется: ушёл — wFault = 0, рампа к
// 40 % от 100 %: 98 % через 1 с.
METHOD PRIVATE PositionerFaultSafePosAction
VAR
    fbTime   : FB_FakeTime;          // подменное время, старт 1 ч
    fbCv     : FB_ControlValve;      // клапан под тестом
    stCmd    : ST_ControlValveCmd;   // команды HMI
    stRetain : ST_DeviceRetain;      // режим Manual по умолчанию
    stCfg    : ST_ControlValveCfg;   // конфигурация (умолчания: 0…100 %, без рампы)
    iStep    : INT;                  // шаг цикла
END_VAR

(* ---- PositionerFaultSafePosAction.method.impl.st ---- *)
coUnit.TEST('ControlValve_PositionerFault_SafePosAction');

stCfg.eFaultAction := E_CvFaultAction.SafePos;
stCfg.rSafePos_pct := 100.0;
stRetain.eRemoteMode := E_DeviceMode.Auto;
fbCv.rPosSpAuto_pct := 40.0;
fbCv(itfTime := fbTime, stCmd := stCmd, stRetain := stRetain, stCfg := stCfg);
stCfg.rRateUp_pctps := 2.0;
stCfg.rRateDown_pctps := 2.0;
fbCv.xPositionerFault := TRUE;
fbTime.Advance(tStep := T#100MS);
fbCv(itfTime := fbTime, stCmd := stCmd, stRetain := stRetain, stCfg := stCfg);
AssertEquals_REAL(Expected := 100.0, Actual := fbCv.rOut_pct, Delta := 0.0, Message := 'safe position at once');
AssertEquals_WORD(Expected := GVL_Const.CV_FLT_POSITIONER, Actual := fbCv.stSts.stCommon.wFault,
                  Message := 'POSITIONER');
AssertTrue(Condition := fbCv.Status = E_Ne107Status.Failure, Message := 'NE 107 Failure');
AssertEquals_WORD(Expected := GVL_Const.CV_STS_SAFE_POS,
                  Actual := fbCv.stSts.stCommon.wStatus AND GVL_Const.CV_STS_SAFE_POS, Message := 'SAFE_POS');
AssertFalse(Condition := fbCv.xAutoActive, Message := 'PID must track');
fbCv.xPositionerFault := FALSE;
// без шага времени
fbCv(itfTime := fbTime, stCmd := stCmd, stRetain := stRetain, stCfg := stCfg);
AssertEquals_WORD(Expected := 0, Actual := fbCv.stSts.stCommon.wFault, Message := 'not latched');
AssertEquals_REAL(Expected := 100.0, Actual := fbCv.rOut_pct, Delta := 0.0,
                  Message := 'ramp starts from safe position');
FOR iStep := 1 TO 10 DO
    fbTime.Advance(tStep := T#100MS);
    fbCv(itfTime := fbTime, stCmd := stCmd, stRetain := stRetain, stCfg := stCfg);
END_FOR
// источник: tools/reference/valve_reference.py, сценарий cv_positioner (100 -> 40, 2 %/s, 1.0 s)
AssertEquals_REAL(Expected := 98.0, Actual := fbCv.rOut_pct, Delta := 1.0E-4, Message := '98 % after 1 s');

coUnit.TEST_FINISHED();

(* ---- RampIndependentOfCycleTime.method.decl.st ---- *)
// Рампа 10 %/с за 2 с даёт одно и то же положение при шаге 10 мс (200 вызовов) и 100 мс (20 вызовов):
// скорость задана в %/с, шаг — фактический ltDt.
METHOD PRIVATE RampIndependentOfCycleTime
VAR
    fbTimeFast   : FB_FakeTime;          // время клапана с шагом 10 мс
    fbTimeSlow   : FB_FakeTime;          // время клапана с шагом 100 мс
    fbFast       : FB_ControlValve;      // клапан, шаг 10 мс
    fbSlow       : FB_ControlValve;      // клапан, шаг 100 мс
    stCmdFast    : ST_ControlValveCmd;   // команды
    stCmdSlow    : ST_ControlValveCmd;   // команды
    stRetainFast : ST_DeviceRetain;      // режим
    stRetainSlow : ST_DeviceRetain;      // режим
    stCfg        : ST_ControlValveCfg;   // рампа 10 %/с
    iStep        : INT;                  // шаг цикла
END_VAR

(* ---- RampIndependentOfCycleTime.method.impl.st ---- *)
coUnit.TEST('ControlValve_Ramp_IndependentOfCycleTime');

stCfg.rRateUp_pctps := 10.0;
stCmdFast.rPosSpMan_pct := 80.0;
stCmdSlow.rPosSpMan_pct := 80.0;
fbFast(itfTime := fbTimeFast, stCmd := stCmdFast, stRetain := stRetainFast, stCfg := stCfg);
fbSlow(itfTime := fbTimeSlow, stCmd := stCmdSlow, stRetain := stRetainSlow, stCfg := stCfg);
FOR iStep := 1 TO 200 DO
    fbTimeFast.Advance(tStep := T#10MS);
    fbFast(itfTime := fbTimeFast, stCmd := stCmdFast, stRetain := stRetainFast, stCfg := stCfg);
END_FOR
FOR iStep := 1 TO 20 DO
    fbTimeSlow.Advance(tStep := T#100MS);
    fbSlow(itfTime := fbTimeSlow, stCmd := stCmdSlow, stRetain := stRetainSlow, stCfg := stCfg);
END_FOR
// источник: tools/reference/valve_reference.py, сценарий cv_cycle_independence: 20.00004 (10 мс) и 20.0 (100 мс)
AssertEquals_REAL(Expected := 20.0, Actual := fbFast.rOut_pct, Delta := 1.0E-4,
                  Message := '10 ms steps: 20 % after 2 s');
AssertEquals_REAL(Expected := 20.0, Actual := fbSlow.rOut_pct, Delta := 1.0E-4,
                  Message := '100 ms steps: 20 % after 2 s');

coUnit.TEST_FINISHED();

(* ---- SlowRamp1msCycleNotStalled.method.decl.st ---- *)
// Рампа 0,003 %/с при цикле 1 мс (CV-14): приращение за шаг 3·10⁻⁶ % меньше половины шага REAL рядом с 70 %
// (7,6·10⁻⁶ %) — в REAL рампа стояла бы на месте. Состояние рампы в LREAL: за 1 с (1000 шагов по 1 мс) выход
// 70,003 % — столько же, сколько при цикле 100 мс (10 шагов). источник: tools/reference/valve_reference.py,
// сценарий cv_slow_ramp.
METHOD PRIVATE SlowRamp1msCycleNotStalled
VAR
    fbTime   : FB_FakeTime;          // подменное время, старт 1 ч
    fbCv     : FB_ControlValve;      // клапан под тестом
    stCmd    : ST_ControlValveCmd;   // команды HMI
    stRetain : ST_DeviceRetain;      // режим Manual по умолчанию
    stCfg    : ST_ControlValveCfg;   // конфигурация (умолчания: 0…100 %, без рампы)

    fbTime2  : FB_FakeTime;          // время второго клапана
    fbCv2    : FB_ControlValve;      // тот же клапан с циклом 100 мс
    stCmd2   : ST_ControlValveCmd;   // его команды
    stRet2   : ST_DeviceRetain;      // его режим
    iStep    : INT;                  // шаг цикла
END_VAR

(* ---- SlowRamp1msCycleNotStalled.method.impl.st ---- *)
coUnit.TEST('ControlValve_SlowRamp1msCycle_NotStalled');

stCmd.rPosSpMan_pct := 70.0;
stCmd2.rPosSpMan_pct := 70.0;
fbCv(itfTime := fbTime, stCmd := stCmd, stRetain := stRetain, stCfg := stCfg);       // Manual, 70 % без рампы
fbCv2(itfTime := fbTime2, stCmd := stCmd2, stRetain := stRet2, stCfg := stCfg);
stCfg.rRateUp_pctps := 0.003;
stCfg.rRateDown_pctps := 0.003;
stCmd.rPosSpMan_pct := 100.0;
stCmd2.rPosSpMan_pct := 100.0;
FOR iStep := 1 TO 1000 DO
    fbTime.AdvanceL(ltStep := LTIME#1MS);
    fbCv(itfTime := fbTime, stCmd := stCmd, stRetain := stRetain, stCfg := stCfg);
END_FOR
FOR iStep := 1 TO 10 DO
    fbTime2.Advance(tStep := T#100MS);
    fbCv2(itfTime := fbTime2, stCmd := stCmd2, stRetain := stRet2, stCfg := stCfg);
END_FOR
AssertEquals_REAL(Expected := 70.003, Actual := fbCv.rOut_pct, Delta := 1.0E-4, Message := '1 ms cycle: ramp moves');
AssertEquals_REAL(Expected := 70.003, Actual := fbCv2.rOut_pct, Delta := 1.0E-4, Message := '100 ms cycle: same');

coUnit.TEST_FINISHED();

(* ---- TightShutBelowThresholdGivesZero.method.decl.st ---- *)
// Плотное закрытие 5 %: задание 4 % — выход 0 % (бит TIGHT_SHUT, 4 мА), 6 % — 6 %. Рампа не залипает под
// порогом: рост 1 %/с, задание 20 %: на 4,5 с выход 0 % (рампа 4,5 %), на 5,0 с ещё 0 % (гистерезис 1 %, CV-13),
// на 6,0 с — 6 %, на 10 с — 10 %.
METHOD PRIVATE TightShutBelowThresholdGivesZero
VAR
    fbTime   : FB_FakeTime;          // подменное время, старт 1 ч
    fbCv     : FB_ControlValve;      // клапан под тестом
    stCmd    : ST_ControlValveCmd;   // команды HMI
    stRetain : ST_DeviceRetain;      // режим Manual по умолчанию
    stCfg    : ST_ControlValveCfg;   // конфигурация (умолчания: 0…100 %, без рампы)
    iStep    : INT;                  // шаг цикла
END_VAR

(* ---- TightShutBelowThresholdGivesZero.method.impl.st ---- *)
coUnit.TEST('ControlValve_TightShut_BelowThresholdGivesZero');

stCfg.rTightShut_pct := 5.0;
stCmd.rPosSpMan_pct := 4.0;
fbCv(itfTime := fbTime, stCmd := stCmd, stRetain := stRetain, stCfg := stCfg);
// источник: tools/reference/valve_reference.py, сценарий cv_tight_ramp (out at sp 4, out at sp 6)
AssertEquals_REAL(Expected := 0.0, Actual := fbCv.rOut_pct, Delta := 0.0, Message := 'below threshold: 0 %');
AssertEquals_WORD(Expected := GVL_Const.CV_STS_TIGHT_SHUT,
                  Actual := fbCv.stSts.stCommon.wStatus AND GVL_Const.CV_STS_TIGHT_SHUT, Message := 'TIGHT_SHUT bit');
AssertEquals_REAL(Expected := 4.0, Actual := fbCv.rOut_mA, Delta := 1.0E-5, Message := '4 mA');
stCmd.rPosSpMan_pct := 6.0;
fbTime.Advance(tStep := T#100MS);
fbCv(itfTime := fbTime, stCmd := stCmd, stRetain := stRetain, stCfg := stCfg);
AssertEquals_REAL(Expected := 6.0, Actual := fbCv.rOut_pct, Delta := 0.0, Message := 'above threshold: as set');
AssertEquals_WORD(Expected := 0, Actual := fbCv.stSts.stCommon.wStatus AND GVL_Const.CV_STS_TIGHT_SHUT,
                  Message := 'no TIGHT_SHUT');
stCfg.rRateUp_pctps := 1.0;
stCmd.rPosSpMan_pct := 0.0;
fbTime.Advance(tStep := T#100MS);
// спад без ограничения — сразу 0
fbCv(itfTime := fbTime, stCmd := stCmd, stRetain := stRetain, stCfg := stCfg);
stCmd.rPosSpMan_pct := 20.0;
FOR iStep := 1 TO 9 DO                                                  // 4,5 с
    fbTime.Advance(tStep := T#500MS);
    fbCv(itfTime := fbTime, stCmd := stCmd, stRetain := stRetain, stCfg := stCfg);
END_FOR
// источник: tools/reference/valve_reference.py, сценарий cv_tight_ramp (out 4.5 s, out 5.0 s, out 10.0 s)
AssertEquals_REAL(Expected := 0.0, Actual := fbCv.rOut_pct, Delta := 0.0, Message := 'ramp 4.5 % below threshold: 0 %');
fbTime.Advance(tStep := T#500MS);
// 5,0 с
fbCv(itfTime := fbTime, stCmd := stCmd, stRetain := stRetain, stCfg := stCfg);
// источник: tools/reference/valve_reference.py, сценарий cv_tight_ramp (out 5.0 s, out 6.0 s); гистерезис CV-13
AssertEquals_REAL(Expected := 0.0, Actual := fbCv.rOut_pct, Delta := 0.0, Message := 'at threshold: still tight shut');
FOR iStep := 11 TO 12 DO                                                // 6,0 с
    fbTime.Advance(tStep := T#500MS);
    fbCv(itfTime := fbTime, stCmd := stCmd, stRetain := stRetain, stCfg := stCfg);
END_FOR
AssertEquals_REAL(Expected := 6.0, Actual := fbCv.rOut_pct, Delta := 1.0E-4, Message := 'released at +1 pct');
FOR iStep := 13 TO 20 DO                                                // 10,0 с
    fbTime.Advance(tStep := T#500MS);
    fbCv(itfTime := fbTime, stCmd := stCmd, stRetain := stRetain, stCfg := stCfg);
END_FOR
AssertEquals_REAL(Expected := 10.0, Actual := fbCv.rOut_pct, Delta := 1.0E-4,
                  Message := 'ramp not stuck under threshold');

coUnit.TEST_FINISHED();

(* ---- TightShutHysteresisNoChatter.method.decl.st ---- *)
// Плотное закрытие 2 % с гистерезисом CV_TIGHT_HYST_PCT = 1 % (CV-13): задание 2,02 %, затем по кругу 1,98 / 2,02 %
// десять вызовов — выход один раз уходит в 0 % и дальше не дёргается; 2,99 % — ещё 0 %; 3,0 % — выход 3,0 %, бит
// TIGHT_SHUT снят.
METHOD PRIVATE TightShutHysteresisNoChatter
VAR
    fbTime   : FB_FakeTime;          // подменное время, старт 1 ч
    fbCv     : FB_ControlValve;      // клапан под тестом
    stCmd    : ST_ControlValveCmd;   // команды HMI
    stRetain : ST_DeviceRetain;      // режим Manual по умолчанию
    stCfg    : ST_ControlValveCfg;   // конфигурация (умолчания: 0…100 %, без рампы)

    iStep    : INT;                  // шаг цикла
    iJumps   : INT;                  // скачков выхода больше 1 %
    rPrev    : REAL;                 // выход прошлого вызова
END_VAR

(* ---- TightShutHysteresisNoChatter.method.impl.st ---- *)
coUnit.TEST('ControlValve_TightShutHysteresis_NoChatter');

stCfg.rTightShut_pct := 2.0;
stRetain.eRemoteMode := E_DeviceMode.Auto;
fbCv.rPosSpAuto_pct := 2.02;
fbCv(itfTime := fbTime, stCmd := stCmd, stRetain := stRetain, stCfg := stCfg);
AssertEquals_REAL(Expected := 2.02, Actual := fbCv.rOut_pct, Delta := 1.0E-4,
                  Message := 'above threshold: no tight shut');
rPrev := fbCv.rOut_pct;
FOR iStep := 1 TO 10 DO
    fbTime.Advance(tStep := T#100MS);
    IF (iStep MOD 2) = 1 THEN
        fbCv.rPosSpAuto_pct := 1.98;
    ELSE
        fbCv.rPosSpAuto_pct := 2.02;
    END_IF
    fbCv(itfTime := fbTime, stCmd := stCmd, stRetain := stRetain, stCfg := stCfg);
    IF ABS(fbCv.rOut_pct - rPrev) > 1.0 THEN
        iJumps := iJumps + 1;
    END_IF
    rPrev := fbCv.rOut_pct;
END_FOR
AssertEquals_INT(Expected := 1, Actual := iJumps, Message := 'one jump into tight shut, no chatter');
AssertEquals_REAL(Expected := 0.0, Actual := fbCv.rOut_pct, Delta := 0.0, Message := 'held in tight shut');
fbCv.rPosSpAuto_pct := 2.99;
fbTime.Advance(tStep := T#100MS);
fbCv(itfTime := fbTime, stCmd := stCmd, stRetain := stRetain, stCfg := stCfg);
AssertEquals_REAL(Expected := 0.0, Actual := fbCv.rOut_pct, Delta := 0.0, Message := 'still tight shut at 2.99 pct');
fbCv.rPosSpAuto_pct := 3.0;
fbTime.Advance(tStep := T#100MS);
fbCv(itfTime := fbTime, stCmd := stCmd, stRetain := stRetain, stCfg := stCfg);
AssertEquals_REAL(Expected := 3.0, Actual := fbCv.rOut_pct, Delta := 1.0E-4,
                  Message := 'released at threshold + hysteresis');
AssertEquals_WORD(Expected := 0, Actual := fbCv.stSts.stCommon.wStatus AND GVL_Const.CV_STS_TIGHT_SHUT,
                  Message := 'TIGHT_SHUT bit cleared');

coUnit.TEST_FINISHED();
